// TIA Portal V20 export
// export: Created 2026-10-20T12:58:39.7495832Z, ExportSetting None, DisplayName Totally Integrated Automation Portal, DisplayVersion V20 Update 6, DisplayName TIA Portal Openness, DisplayVersion V20 Update 6, DisplayName TIA Portal Version Control Interface, DisplayVersion V20 Update 6, DisplayName SINAMICS Startdrive Advanced, DisplayVersion V20 SP1, DisplayName SINAMICS Startdrive G130, G150, S120, S150, SINAMICS MV, G220, S200, S210, DisplayVersion V20 SP1, DisplayName SINAMICS Startdrive G110M, G120, G120C, G120D, G120P, G115D, DisplayVersion V20 SP1, DisplayName STEP 7 Professional, DisplayVersion V20 Update 6, DisplayName STEP 7 Safety, DisplayVersion V20 Update 2, DisplayName WinCC Basic/Comfort/Advanced, DisplayVersion V20 Update 6, DisplayName WinCC Unified, DisplayVersion V20 Update 6
VAR_GLOBAL   // PLC tag table "Default table"
   System_Byte AT %MB1159 : Byte;
   FirstScan AT %M1159.0 : Bool;
   DiagStatusUpdate AT %M1159.1 : Bool;
   AlwaysTRUE AT %M1159.2 : Bool;
   AlwaysFALSE AT %M1159.3 : Bool;
   Clock_Byte AT %MB1160 : Byte;
   Clock_10Hz AT %M1160.0 : Bool;
   Clock_5Hz AT %M1160.1 : Bool;
   "Clock_2.5Hz" AT %M1160.2 : Bool;
   Clock_2Hz AT %M1160.3 : Bool;
   "Clock_1.25Hz" AT %M1160.4 : Bool;
   Clock_1Hz AT %M1160.5 : Bool;
   "Clock_0.625Hz" AT %M1160.6 : Bool;
   "Clock_0.5Hz" AT %M1160.7 : Bool;
   "System_Byte(1)" AT %MB1 : Byte;
   Tag_1 AT %M2000.0 : Bool;
   Tag_2 AT %M2000.1 : Bool;
   Tag_3 AT %M2000.2 : Bool;
   Reintegration AT %M2000.3 : Bool;
   Error_Word_1 AT %MW2001 : Word;
   "Auto_Start_Lector(4)" AT %M20.4 : Bool;
   "Auto_Stop_Lector(4)" AT %M25.2 : Bool;
   "Auto_Stop_Lector(1)" AT %M20.6 : Bool;
   "Auto_Stop_Lector(2)" AT %M20.7 : Bool;
   "Auto_Start_Lector(1)" AT %M19.6 : Bool;
   "Auto_Start_Lector(2)" AT %M20.2 : Bool;
   "Auto_Stop_Lector(3)" AT %M25.1 : Bool;
   "Auto_Stop_Lector(5)" AT %M25.3 : Bool;
   "Auto_Start_Lector(5)" AT %M20.5 : Bool;
   "Auto_Start_Lector(3)" AT %M20.3 : Bool;
   Force_System_1 AT %M25.5 : Bool;
   VTD_System_Selected_HMI AT %MW1234 : UInt;
   Initialization AT %M19.4 : Bool;
   Save_Settings AT %M0.1 : Bool;
   "LE_Bypass(1)" AT %M704.1 : Bool;
   "LE_Bypass(4)" AT %M704.4 : Bool;
   "LE_Bypass(5)" AT %M704.5 : Bool;
   "LE_Bypass(2)" AT %M704.2 : Bool;
   "LE_Bypass(3)" AT %M704.3 : Bool;
   Reset_Comissioning AT %M70.0 : Bool;
   "Clear_OT(1)" AT %M154.4 : Bool;
   "Clear_OT(2)" AT %M154.5 : Bool;
   "Clear_OT(4)" AT %M154.7 : Bool;
   "Clear_OT(3)" AT %M154.6 : Bool;
   "Clear_OT(5)" AT %M155.0 : Bool;
   System_3_Busy AT %M39.7 : Bool;
   System_4_Busy AT %M60.2 : Bool;
   System_5_Busy AT %M60.3 : Bool;
   System_2_Busy AT %M39.6 : Bool;
   System_1_Busy AT %M19.5 : Bool;
   L3_OK AT %M39.4 : Bool;
   L4_OK AT %M39.0 : Bool;
   L8_OK AT %M39.5 : Bool;
   L5_OK AT %M39.1 : Bool;
   L1_OK AT %M26.6 : Bool;
   L2_OK AT %M26.7 : Bool;
   L7_OK AT %M39.3 : Bool;
   L6_OK AT %M39.2 : Bool;
   L7_Estop AT %M71.0 : Bool;
   L1_Estop AT %M61.6 : Bool;
   L6_Estop AT %M70.6 : Bool;
   L8_Estop AT %M71.1 : Bool;
   L2_Estop AT %M61.7 : Bool;
   L5_Estop AT %M70.4 : Bool;
   L4_Estop AT %M70.3 : Bool;
   L3_Estop AT %M70.2 : Bool;
   LGX_Secure_Access_2 AT %M71.5 : Bool;
   LGX_Secure_Access_3 AT %M71.6 : Bool;
   LGX_Secure_Access_1 AT %M71.4 : Bool;
   LGX_ReadyToReceive_3 AT %M71.3 : Bool;
   LGX_ReadyToReceive_2 AT %M71.2 : Bool;
   LGX_ReadyToReceive_1 AT %M61.5 : Bool;
   Dbug AT %M71.7 : Bool;
   Reset_Locks AT %M80.2 : Bool;
   HMI_2_Local_Mode AT %M80.5 : Bool;
   Comissioning_Var AT %M80.6 : Bool;
   Material_Selection_O_3 AT %M82.1 : Bool;
   MR_O_2 AT %M82.0 : Bool;
   Material_Selection_I_3 AT %M81.3 : Bool;
   MR_O_1 AT %M81.6 : Bool;
   MR_Delay_O AT %MD200 : Time;
   MR_I_1 AT %M81.0 : Bool;
   MR_Delay_I AT %MD196 : Time;
   Material_Selection_I_2 AT %M81.1 : Bool;
   Material_Selection_O_2 AT %M81.7 : Bool;
   Material_Selection_I_1 AT %M80.7 : Bool;
   MR_O_3 AT %M82.2 : Bool;
   MR_I_3 AT %M81.4 : Bool;
   Material_Selection_O_1 AT %M81.5 : Bool;
   MR_I_2 AT %M81.2 : Bool;
   Starting_Pallet_1 AT %M102.1 : Bool;
   Starting_Pallet_2 AT %M102.2 : Bool;
   Starting_Pallet_3 AT %M102.3 : Bool;
   Time_1_end_Ecnv AT %MD232 : Time;
   Time_2_Start_Ecnv AT %MD236 : Time;
   Time_3_Ecnv AT %MD244 : Time;
   Time_1_end_Buffers AT %MD208 : Time;
   Time_2_Start_Buffers AT %MD212 : Time;
   Time_1_Start_Ecnv AT %MD228 : Time;
   Time_3_Buffers AT %MD224 : Time;
   Time_2_End_Ecnv AT %MD240 : Time;
   Time_2_End_Buffers AT %MD220 : Time;
   Time_1_Start_Buffers AT %MD204 : Time;
END_VAR
